Fanuc KAREL source: kb00124.KL

PROGRAM KB00124
%STACKSIZE=65535
%PRIORITY=65535
%NOLOCKGROUP
VAR
P1 : STRING[80]
P2 : INTEGER
BEGIN
P1='A'
P2=1
MSG_CONNECT(P1,P2)
END KB00124
